Universal Robots URScript: T014_zai-org_GLM-4.7-FP8_edit_perf_rep1.urscript

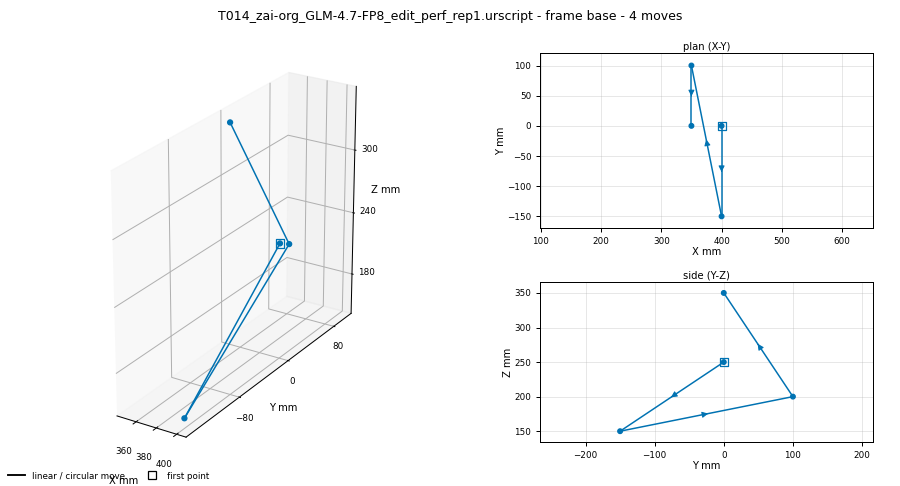
[picture p0: tool path of T014_zai-org_GLM-4.7-FP8_edit_perf_rep1.urscript in frame base, 4 of 6 moves have a stored position in this frame; points joined in program order, loops and branches not executed]
# Task: T014 — Hybrid multi-angle camera inspection (Optimized)
# Generated by ENFIELD IR→URScript Translator
# Operating mode: hybrid | Max TCP speed: 0.200 m/s
# Robot: ur5e
#
# WARNING: This is auto-generated code for SIMULATION ONLY.
# Do NOT deploy to a physical robot without safety review.

def task_T014():
  # [0] E-Stop verify
  # E-Stop safety check (hardware-enforced on UR controller)
  if (get_digital_in(0) == True):
    popup("E-Stop active — aborting program.", error=True)
    halt
  end

  # [1] Home (Increased joint velocity/acceleration for faster reset)
  movej([0.0000, -1.5708, 1.5708, -1.5708, -1.5708, 0.0000], a=2.0000, v=1.5000)

  # [2] Top-down view position (Max TCP speed, higher accel, zero radius for precision)
  movel(p[0.400000, 0.000000, 0.250000, 0.0000, 3.1416, 0.0000], a=1.2000, v=0.2000, r=0.0000)

  # [3] Camera trigger ON
  set_digital_out(2, True)

  # [4] Capture top view (Reduced sleep time for faster cycle)
  sleep(0.1000)

  # [5] Camera trigger OFF
  set_digital_out(2, False)

  # [6] Side view position (Max TCP speed, higher accel, zero radius)
  movel(p[0.400000, -0.150000, 0.150000, 0.0000, 3.1416, 0.0000], a=1.2000, v=0.2000, r=0.0000)

  # [7] Camera trigger ON
  set_digital_out(2, True)

  # [8] Capture side view (Reduced sleep time)
  sleep(0.1000)

  # [9] Camera trigger OFF
  set_digital_out(2, False)

  # [10] Angled view position (Max TCP speed, higher accel, zero radius)
  movel(p[0.350000, 0.100000, 0.200000, 0.0000, 3.1416, 0.0000], a=1.2000, v=0.2000, r=0.0000)

  # [11] Camera trigger ON
  set_digital_out(2, True)

  # [12] Capture angled view (Reduced sleep time)
  sleep(0.1000)

  # [13] Camera trigger OFF
  set_digital_out(2, False)

  # [14] Retract (Max speed, blend allowed as no inspection occurs here)
  movel(p[0.350000, 0.000000, 0.350000, 0.0000, 3.1416, 0.0000], a=1.2000, v=0.2000, r=0.0500)

  # [15] Return home (Increased joint velocity/acceleration)
  movej([0.0000, -1.5708, 1.5708, -1.5708, -1.5708, 0.0000], a=2.0000, v=1.5000)

end

# Entry point
task_T014()
